(* IEC 61131-3 sources: ia2/library/process-control/pous (part 2) *)

(* ---- fb_pid_3step.st ---- *)
(*
  FB_PID_3STEP — step (3-step) PID: open/close pulse control of a motorized actuator,
  supporting both no-position-feedback (travel-time integral estimate) and
  with-feedback wiring.

  ~ Standard step PID / 3-step output controller (step controller / 3-step PID, driving
  integrating-type actuators such as motorized control valves and motorized dampers),
  found in every major DCS/PLC standard library.

  Purpose: closed-loop control of a motorized actuator (motorized valve / motorized
  damper, which is itself an integrating element: energized it runs open/close, de-energized
  it stops in place). Without a position transmitter, estimate position by integrating
  travel time (pos_fb < 0); with a 4-20 mA position feedback, use it directly.

  Behavior:
    1) Position estimate pos_est: pos_fb >= 0 takes the feedback directly (clamped
       0..100); otherwise integrate from the previous scan's output and the travel time:
       an open pulse adds +100*dt_s/motor_time_s, a close pulse decrements likewise
       (clamped 0..100).
    2) An internal positional PID (reverse-acting e = sp - pv, D on PV with automatic
       3*dt_s PT1 filtering) computes the target position target 0..100; integral
       back-calculation anti-windup; in manual, target tracks pos_est so the return to
       auto is bumpless. For direct-acting scenarios, invert pv/sp externally.
    3) Three-step output: position deviation = target - pos_est;
       > deadband_pct emits an open pulse, < -deadband_pct emits a close pulse, within
       the deadband stop. In auto, once a pulse is emitted it is held at least
       min_pulse_s (to avoid short pulses hammering the contactor); manual jogs
       man_open/man_close pass through (no minimum pulse width, mutually interlocked
       when both are commanded), constrained only by the travel limits. A reversal must
       pass through one scan fully stopped (stop before reversing). At a travel boundary
       (pos_est reaching 0 or 100), stop that direction's pulse immediately.
    Tuning tip: deadband_pct should be larger than the travel corresponding to the
    minimum pulse width (min_pulse_s / motor_time_s * 100%), otherwise it will still
    overshoot and oscillate within the deadband.

  Inputs:
    pv           REAL  process value
    sp           REAL  setpoint
    kp           REAL  proportional gain
    ti_s         REAL  integral time s (0 = no integral)
    td_s         REAL  derivative time s (0 = derivative off)
    dt_s         REAL  sample period s (<= 0 holds this scan, no action)
    motor_time_s REAL  actuator full-travel time s (0->100%; used for estimation and limits)
    min_pulse_s  REAL  minimum pulse width in auto s
    deadband_pct REAL  position deadband % (no action within the deviation deadband)
    auto         BOOL  TRUE auto / FALSE manual jog
    man_open     BOOL  manual open jog (interlocked, no action when commanded with man_close)
    man_close    BOOL  manual close jog
    pos_fb       REAL  position feedback 0..100 % (< 0 = no feedback, use travel estimate)
  Outputs:
    q_open  BOOL  open-direction pulse output
    q_close BOOL  close-direction pulse output
    pos_est REAL  position estimate/feedback 0..100 %
*)
FUNCTION_BLOCK FB_PID_3STEP
  VAR_INPUT
    pv           : REAL;
    sp           : REAL;
    kp           : REAL := 1.0;
    ti_s         : REAL := 0.0;
    td_s         : REAL := 0.0;
    dt_s         : REAL := 0.1;
    motor_time_s : REAL := 60.0;
    min_pulse_s  : REAL := 0.5;
    deadband_pct : REAL := 1.0;
    auto         : BOOL := TRUE;
    man_open     : BOOL := FALSE;
    man_close    : BOOL := FALSE;
    pos_fb       : REAL := -1.0;
  END_VAR
  VAR_OUTPUT
    q_open  : BOOL;
    q_close : BOOL;
    pos_est : REAL;
  END_VAR
  VAR
    i_acc     : REAL; (* positional-PID integral term (back-calculation bumpless) *)
    pv_f      : REAL; (* D-term PT1 filter state *)
    pv_f_prev : REAL;
    t_f       : REAL;
    e         : REAL;
    p_term    : REAL;
    d_term    : REAL;
    target    : REAL; (* PID target position 0..100 *)
    err_pos   : REAL; (* position deviation target - pos_est *)
    pulse_t   : REAL; (* elapsed duration of the current pulse s *)
    open_req  : BOOL; (* open-direction demand this scan *)
    close_req : BOOL;
    init_done : BOOL; (* filter-state first-scan alignment flag *)
  END_VAR

  IF dt_s <= 0.0 THEN
    RETURN; (* invalid sample period: hold *)
  END_IF;

  IF NOT init_done THEN
    pv_f := pv;
    pv_f_prev := pv;
    init_done := TRUE;
  END_IF;

  (* 1) Position estimate: use feedback directly when available; otherwise integrate from the previous scan's output over the travel time *)
  IF pos_fb >= 0.0 THEN
    pos_est := pos_fb;
  ELSE
    IF motor_time_s > 0.0 THEN
      IF q_open THEN
        pos_est := pos_est + 100.0 * dt_s / motor_time_s;
      END_IF;
      IF q_close THEN
        pos_est := pos_est - 100.0 * dt_s / motor_time_s;
      END_IF;
    END_IF;
  END_IF;
  IF pos_est > 100.0 THEN
    pos_est := 100.0;
  ELSIF pos_est < 0.0 THEN
    pos_est := 0.0;
  END_IF;

  (* 2) Positional PID -> target position (reverse-acting; D on PV, automatic 3*dt_s filtering) *)
  t_f := 3.0 * dt_s;
  pv_f := pv_f + dt_s / (t_f + dt_s) * (pv - pv_f);
  e := sp - pv;
  p_term := kp * e;
  d_term := 0.0;
  IF td_s > 0.0 THEN
    d_term := 0.0 - kp * td_s * (pv_f - pv_f_prev) / dt_s;
  END_IF;
  pv_f_prev := pv_f;

  IF auto THEN
    IF ti_s > 0.0 THEN
      i_acc := i_acc + kp * dt_s / ti_s * e;
    END_IF;
    target := p_term + i_acc + d_term;
  ELSE
    target := pos_est; (* Manual: target tracks the current position, bumpless return to auto *)
  END_IF;
  IF target > 100.0 THEN
    target := 100.0;
  ELSIF target < 0.0 THEN
    target := 0.0;
  END_IF;
  IF ti_s > 0.0 OR NOT auto THEN
    i_acc := target - p_term - d_term; (* Back-calculation: anti-windup + bumpless *)
  END_IF;

  (* 3) Three-step output demand *)
  IF auto THEN
    err_pos := target - pos_est;
    open_req := err_pos > deadband_pct;
    close_req := err_pos < 0.0 - deadband_pct;
  ELSE
    open_req := man_open AND NOT man_close; (* Manual jog passes through, interlocked when both commanded *)
    close_req := man_close AND NOT man_open;
  END_IF;

  (* Travel limits: at a boundary, stop emitting that direction's pulse (same in manual/auto) *)
  IF pos_est >= 100.0 THEN
    open_req := FALSE;
  END_IF;
  IF pos_est <= 0.0 THEN
    close_req := FALSE;
  END_IF;

  (* Pulse timing and output: in auto, dropping the demand must satisfy the minimum
     pulse width; in manual, dropping stops immediately; a reversal must pass through
     one scan fully stopped (the current direction drops first, the reverse is allowed
     only on the next scan) *)
  IF q_open OR q_close THEN
    pulse_t := pulse_t + dt_s;
  END_IF;

  IF q_open THEN
    IF pos_est >= 100.0 THEN
      q_open := FALSE; (* at limit, stop *)
    ELSIF NOT open_req AND (NOT auto OR pulse_t >= min_pulse_s) THEN
      q_open := FALSE;
    END_IF;
  ELSIF q_close THEN
    IF pos_est <= 0.0 THEN
      q_close := FALSE;
    ELSIF NOT close_req AND (NOT auto OR pulse_t >= min_pulse_s) THEN
      q_close := FALSE;
    END_IF;
  ELSE
    pulse_t := 0.0;
    IF open_req THEN
      q_open := TRUE;
    ELSIF close_req THEN
      q_close := TRUE;
    END_IF;
  END_IF;
END_FUNCTION_BLOCK

(* ---- fb_pid_pos.st ---- *)
(*
  FB_PID_POS — positional (absolute-output) PID controller with observable p/i/d terms,
  SP weighting, derivative-on-PV (D on PV + PT1 filter), back-calculation anti-windup
  and bumpless transfer.

  ~ Standard positional PID (absolute-output form, observable P/I/D terms, SP weighting
  b, derivative acting on PV), found in every major DCS/PLC standard library.

  Purpose: complements the velocity-form FB_PID -- for loops that need to observe/debug
  the integral term, want SP weighting (b < 1 suppresses the proportional kick on a
  setpoint step), or need an absolute-quantity output downstream. For incremental
  output / cascade relay scenarios, FB_PID is still recommended.

  Algorithm (positional):
    e   := sp - pv (reverse-acting, default); direct = TRUE gives e := pv - sp
    e_p := b*sp - pv (the SP-weighted deviation used only by the P term; reversed when direct)
    p_part := kp * e_p
    i_part := i_part + kp*dt_s/ti_s * e (accumulated when ti_s > 0)
    d_part := -kp*td_s * d(pv_f)/dt (derivative acts on PV: no kick on an SP step;
              pv first passes a PT1 filter, t_dfilt_s <= 0 takes 3*dt_s automatically;
              sign goes positive when direct)
    out := p_part + i_part + d_part + ff, clamped to [out_min, out_max]
  Anti-windup and bumpless (back-calculation): each scan wraps up by back-calculating i_part as
    i_part := out - p_part - d_part - ff
  -- on clamping the integral is pulled back (no windup); in manual/track the output
  follows the supplied value and i_part back-calculates in step, so the return to auto
  has no jump. When ti_s = 0 (no integral), i_part is back-calculated only during
  manual/track (where it is a fixed bias / manual-reset term, not overwritten by
  clamping events during auto, keeping the offset characteristic of P-type control
  stable).
  Mode priority: track > NOT auto (manual) > auto (same as FB_PID).
  Identity: in every mode out = p_part + i_part + d_part + ff (after clamping, except
  on an auto clamping scan with ti_s = 0) -- the sum of the terms is the output,
  intuitive for debugging.

  Inputs:
    pv          REAL  process value
    sp          REAL  setpoint
    kp          REAL  proportional gain
    ti_s        REAL  integral time s (0 = no integral)
    td_s        REAL  derivative time s (0 = derivative off)
    t_dfilt_s   REAL  derivative pre-filter PT1 time constant s (<= 0 = auto 3*dt_s)
    sp_weight_b REAL  SP weighting coefficient b (acts on the P term only; 1 = no weighting,
                      0 = the P term sees pv only -- an SP step gives no proportional kick at all)
    dt_s        REAL  sample period s (<= 0 holds this scan, no action)
    direct      BOOL  TRUE = direct-acting (pv up -> out up), FALSE = reverse-acting
    auto        BOOL  TRUE auto / FALSE manual
    manual_out  REAL  manual output value
    out_min     REAL  output low limit (assumes out_min < out_max)
    out_max     REAL  output high limit
    ff          REAL  feedforward (added to output before clamp)
    track       BOOL  output-tracking enable (highest priority)
    track_value REAL  tracking value
  Outputs:
    out    REAL  control output (clamped in every mode)
    dev    REAL  deviation (reverse-acting sp-pv / direct-acting pv-sp, without SP weighting)
    p_part REAL  proportional term (includes SP weighting)
    i_part REAL  integral term (includes back-calculation correction)
    d_part REAL  derivative term
*)
FUNCTION_BLOCK FB_PID_POS
  VAR_INPUT
    pv          : REAL;
    sp          : REAL;
    kp          : REAL := 1.0;
    ti_s        : REAL := 0.0;
    td_s        : REAL := 0.0;
    t_dfilt_s   : REAL := 0.0;
    sp_weight_b : REAL := 1.0;
    dt_s        : REAL := 0.1;
    direct      : BOOL := FALSE;
    auto        : BOOL := TRUE;
    manual_out  : REAL := 0.0;
    out_min     : REAL := 0.0;
    out_max     : REAL := 100.0;
    ff          : REAL := 0.0;
    track       : BOOL := FALSE;
    track_value : REAL := 0.0;
  END_VAR
  VAR_OUTPUT
    out    : REAL;
    dev    : REAL;
    p_part : REAL;
    i_part : REAL;
    d_part : REAL;
  END_VAR
  VAR
    pv_f      : REAL; (* PV after the D-term PT1 filter *)
    pv_f_prev : REAL; (* previous-scan filtered value, for the backward difference *)
    t_f       : REAL; (* filter time constant actually used *)
    d_pv      : REAL; (* rate of change of the filtered PV, units/s *)
    e         : REAL; (* control deviation (includes the action direction) *)
    e_p       : REAL; (* P-term deviation (SP weighting b) *)
    init_done : BOOL; (* filter-state first-scan alignment flag *)
  END_VAR

  IF dt_s <= 0.0 THEN
    RETURN; (* invalid sample period: hold output and history unchanged *)
  END_IF;

  IF NOT init_done THEN
    pv_f := pv; (* align the filter state: no spurious startup derivative *)
    pv_f_prev := pv;
    init_done := TRUE;
  END_IF;

  (* D-term pre-filter PT1 + backward difference (same core as FB_DERIV) *)
  t_f := t_dfilt_s;
  IF t_f <= 0.0 THEN
    t_f := 3.0 * dt_s;
  END_IF;
  pv_f := pv_f + dt_s / (t_f + dt_s) * (pv - pv_f);
  d_pv := (pv_f - pv_f_prev) / dt_s;
  pv_f_prev := pv_f;

  (* Deviation (by action direction) and the SP-weighted P deviation *)
  IF direct THEN
    e := pv - sp;
    e_p := pv - sp_weight_b * sp;
  ELSE
    e := sp - pv;
    e_p := sp_weight_b * sp - pv;
  END_IF;
  dev := e;

  p_part := kp * e_p;

  d_part := 0.0;
  IF td_s > 0.0 THEN
    (* Derivative acts on PV (no kick on an SP step): reverse-acting, rising pv should push the output down -> negative sign *)
    IF direct THEN
      d_part := kp * td_s * d_pv;
    ELSE
      d_part := 0.0 - kp * td_s * d_pv;
    END_IF;
  END_IF;

  IF track THEN
    (* Output tracking: follows track_value unconditionally, highest priority *)
    out := track_value;
  ELSIF NOT auto THEN
    (* Manual: follows manual_out; the i_part back-calculation guarantees a bumpless return to auto *)
    out := manual_out;
  ELSE
    IF ti_s > 0.0 THEN
      i_part := i_part + kp * dt_s / ti_s * e;
    END_IF;
    out := p_part + i_part + d_part + ff;
  END_IF;

  (* Output clamp *)
  IF out > out_max THEN
    out := out_max;
  ELSIF out < out_min THEN
    out := out_min;
  END_IF;

  (* Back-calculate i_part: makes P+I+D+ff always equal the clamped output -> clamping
     gives anti-windup and manual/track gives bumpless alignment. When ti_s = 0,
     back-calculate only during manual/track (see header note) *)
  IF ti_s > 0.0 OR track OR NOT auto THEN
    i_part := out - p_part - d_part - ff;
  END_IF;
END_FUNCTION_BLOCK

(* ---- fb_pulser.st ---- *)
(*
  FB_PULSER — periodic pulse generator.

  Purpose: periodic air-cannon / air-hammer silo purging, periodic lubrication, heartbeat output.
  Example: once enabled, output a pulse_len_s-wide pulse every period_s seconds (the pulse comes at the period start).

  Behavior:
    while enabled, the phase phase_s accumulates by dt_s manually; q := TRUE while
    phase_s < pulse_len_s, wrapping at period_s (subtraction wrap, so the long-term
    cadence does not drift).
    NOT enable or invalid parameters (period_s/dt_s <= 0) -> q := FALSE and phase cleared
    (re-enabling starts from the pulse).
    pulse_len_s >= period_s -> q is always TRUE (continuous output by definition).

  Inputs:
    enable      BOOL  enable
    period_s    REAL  pulse period s
    pulse_len_s REAL  pulse width s
    dt_s        REAL  sample period s
  Outputs:
    q BOOL  pulse output
*)
FUNCTION_BLOCK FB_PULSER
  VAR_INPUT
    enable      : BOOL;
    period_s    : REAL := 60.0;
    pulse_len_s : REAL := 1.0;
    dt_s        : REAL := 0.1;
  END_VAR
  VAR_OUTPUT
    q : BOOL;
  END_VAR
  VAR
    phase_s : REAL; (* phase within the period 0..period_s, manual timing in place of TP/TON *)
  END_VAR

  IF NOT enable OR period_s <= 0.0 OR dt_s <= 0.0 THEN
    phase_s := 0.0;
    q := FALSE;
    RETURN;
  END_IF;

  (* Emit the pulse by the current phase first (TRUE immediately on the first enabled period), then advance the phase *)
  q := phase_s < pulse_len_s;

  phase_s := phase_s + dt_s;
  IF phase_s >= period_s THEN
    phase_s := phase_s - period_s; (* subtraction wrap, keeps the long-term cadence *)
  END_IF;
END_FUNCTION_BLOCK

(* ---- fb_pv_hold.st ---- *)
(*
  FB_PV_HOLD — bad-PV hold / substitute.

  ~ Standard bad-value handling block (last-good hold / substitute value, including
  bad-value timeout degradation), the standard line of defense before a measurement
  enters a control loop; every major DCS/PLC input-processing chain has an equivalent
  mechanism.

  Purpose: on transmitter open-circuit/over-range (e.g. FB_SCALE.fault, or the inverse
  of FB_MID3.q_fail used as good), give the downstream loop a controlled PV: hold the
  last good value first to ride out chatter, then on timeout hold/substitute/follow as
  configured, while emitting q_bad/q_timeout for alarming and loop-to-manual logic.

  Behavior:
    good = TRUE: out := u, remember the last good value, clear q_bad/q_timeout, clear
    the bad-value timer.
    good = FALSE: q_bad := TRUE, accumulate the bad-value timer (manual dt_s):
      before timeout_s: out := last good value (short chatter rides through on hold);
      at timeout_s (timeout_s = 0 immediately): q_timeout := TRUE, then by mode:
        mode = 0: keep holding the last good value;
        mode = 1: out := sub_value (substitute value, e.g. a safe-side setting);
        mode = 2: out := u (follow the raw value -- just raise the alarm flag without
                  intervening, downstream handles it).
    When bad on the very first scan, the last good value takes the current u (no better history).
    dt_s <= 0 -> the bad-value timer does not advance (when timeout_s > 0, the hold segment is maintained).

  Inputs:
    u         REAL  input (raw PV)
    good      BOOL  input valid (FALSE = bad value; feed the inverse of a quality bit / open-circuit decision)
    mode      REAL  0 = hold last good value / 1 = substitute value / 2 = follow raw value
    sub_value REAL  substitute value (used by mode = 1)
    timeout_s REAL  bad-value persistence timeout s (0 = act by mode immediately; > 0 hold first)
    dt_s      REAL  sample period s
  Outputs:
    out       REAL  processed PV
    q_bad     BOOL  in bad value (level)
    q_timeout BOOL  bad value has timed out (mode in effect)
*)
FUNCTION_BLOCK FB_PV_HOLD
  VAR_INPUT
    u         : REAL;
    good      : BOOL := TRUE;
    mode      : REAL := 0.0;
    sub_value : REAL := 0.0;
    timeout_s : REAL := 0.0;
    dt_s      : REAL := 0.1;
  END_VAR
  VAR_OUTPUT
    out       : REAL;
    q_bad     : BOOL;
    q_timeout : BOOL;
  END_VAR
  VAR
    last_good : REAL; (* last good value *)
    bad_t     : REAL; (* bad-value accumulated persistence time s *)
    init_done : BOOL; (* first-scan seeding flag *)
  END_VAR

  IF NOT init_done THEN
    last_good := u; (* even when bad on the first scan, take the current u as the held value *)
    init_done := TRUE;
  END_IF;

  IF good THEN
    last_good := u;
    out := u;
    q_bad := FALSE;
    q_timeout := FALSE;
    bad_t := 0.0;
    RETURN;
  END_IF;

  q_bad := TRUE;

  (* Before timeout: hold the last good value (the segment that rides out short chatter) *)
  IF timeout_s > 0.0 THEN
    IF dt_s > 0.0 THEN
      bad_t := bad_t + dt_s;
    END_IF;
    IF bad_t < timeout_s THEN
      out := last_good;
      q_timeout := FALSE;
      RETURN;
    END_IF;
  END_IF;

  (* On timeout (or immediately when timeout_s = 0): act by mode *)
  q_timeout := TRUE;
  IF mode >= 1.5 THEN
    out := u;         (* 2 = follow raw value *)
  ELSIF mode >= 0.5 THEN
    out := sub_value; (* 1 = substitute value *)
  ELSE
    out := last_good; (* 0 = hold last good value *)
  END_IF;
END_FUNCTION_BLOCK

(* ---- fb_pwm.st ---- *)
(*
  FB_PWM — time-proportioning output (0..100% command -> fixed-period duty-cycle on/off).

  ~ Time-proportioning (time-proportioning / PWM): continuous quantity -> periodic
  on/off, the customary form for solid-state-relay / solenoid-valve temperature control.

  Purpose: a PID output driving an on/off actuator via a solid-state relay / solenoid
  valve: electric heaters, steam on/off valves, dosing pumps.
  Behavior:
    Phase accumulator as in FB_PULSER: phase_s accumulates by dt_s, wraps by subtraction
    at period_s (so the long-term cadence does not drift); q := phase_s < on_s.
    on_s := u/100 * period_s (u clamped 0..100 first).
    Minimum on/off times (protecting the contactor/SSR/valve, implemented by clamping the effective duty):
      0 < on_s < min_on_s            -> on_s raised to min_on_s;
      0 < period_s - on_s < min_off_s -> on_s squeezed to period_s - min_off_s
      (the off side has higher priority; if min_on_s + min_off_s > period_s the
      parameters are contradictory and the off side wins -- at the extreme it stays
      permanently off, so do not tune it this way).
    u <= 0 -> off for the whole period; u >= 100 -> on for the whole period (full scale
    is unaffected by the minimum on/off clamp).
    NOT enable or period_s/dt_s <= 0 -> q := FALSE and phase cleared (re-enabling starts
    from the period start, on first then off).
    A change in u takes effect immediately (the comparison threshold within the period
    changes at once, no need to wait for the next period).

  Inputs:
    u         REAL  command 0..100 %
    period_s  REAL  PWM period s
    min_on_s  REAL  minimum on time s (0 = no limit)
    min_off_s REAL  minimum off time s (0 = no limit)
    enable    BOOL  enable
    dt_s      REAL  sample period s
  Outputs:
    q         BOOL  time-proportioning output
*)
FUNCTION_BLOCK FB_PWM
  VAR_INPUT
    u         : REAL;
    period_s  : REAL := 10.0;
    min_on_s  : REAL := 0.0;
    min_off_s : REAL := 0.0;
    enable    : BOOL;
    dt_s      : REAL := 0.1;
  END_VAR
  VAR_OUTPUT
    q : BOOL;
  END_VAR
  VAR
    phase_s : REAL; (* phase within the period, manual timing in place of TP/TON *)
    uc      : REAL;
    on_s    : REAL; (* effective on-duration this scan *)
    off_s   : REAL;
  END_VAR

  IF NOT enable OR period_s <= 0.0 OR dt_s <= 0.0 THEN
    phase_s := 0.0;
    q := FALSE;
    RETURN;
  END_IF;

  uc := u;
  IF uc < 0.0 THEN
    uc := 0.0;
  ELSIF uc > 100.0 THEN
    uc := 100.0;
  END_IF;

  on_s := uc * period_s / 100.0;

  (* Minimum on: raise the effective duty (u=0 unaffected) *)
  IF on_s > 0.0 AND on_s < min_on_s THEN
    on_s := min_on_s;
  END_IF;

  (* Minimum off: lower the effective duty (at u=100, off=0 so it does not trigger, stays permanently on) *)
  off_s := period_s - on_s;
  IF off_s > 0.0 AND off_s < min_off_s THEN
    on_s := period_s - min_off_s;
    IF on_s < 0.0 THEN
      on_s := 0.0;
    END_IF;
  END_IF;

  q := phase_s < on_s;

  phase_s := phase_s + dt_s;
  IF phase_s >= period_s THEN
    phase_s := phase_s - period_s; (* subtraction wrap, keeps the long-term cadence *)
  END_IF;
END_FUNCTION_BLOCK

(* ---- fb_ramp.st ---- *)
(*
  FB_RAMP — setpoint ramp generator (rate-limited approach to a fixed target).

  ~ Standard setpoint ramp generator.

  Purpose: gentle setpoint changes (avoiding step shocks to actuators/process),
  segmented heat-up/pressure-up curves.
  Difference from FB_RATE_LIMIT: this block moves toward a fixed target and reports
  ramping; RATE_LIMIT continuously follows a changing input and only clamps the
  per-second change.

  Behavior:
    out approaches target at rate_up (upward) / rate_dn (downward, supplied positive)
    units per second, and on arrival ramping := FALSE. A rate of 0 means a direct
    step in that direction.
    track level-active: out follows track_value unconditionally and ramping := FALSE;
    after track is released, the ramp continues from the current value toward target
    (the bumpless-startup idiom: track-align to the current process value first, then
    release to start ramping).
    dt_s <= 0 -> hold. Note out initializes to 0: on the first startup scan, prefer
    aligning with track.

  Inputs:
    target      REAL  target value
    rate_up     REAL  upward rate units/s (0 = step)
    rate_dn     REAL  downward rate units/s (supplied positive; 0 = step)
    dt_s        REAL  sample period s
    track       BOOL  tracking enable (level-active)
    track_value REAL  tracking value
  Outputs:
    out     REAL  ramp output
    ramping BOOL  ramp in progress (target not yet reached)
*)
FUNCTION_BLOCK FB_RAMP
  VAR_INPUT
    target      : REAL;
    rate_up     : REAL := 0.0;
    rate_dn     : REAL := 0.0;
    dt_s        : REAL := 0.1;
    track       : BOOL := FALSE;
    track_value : REAL := 0.0;
  END_VAR
  VAR_OUTPUT
    out     : REAL;
    ramping : BOOL;
  END_VAR
  VAR
    delta : REAL;
    step  : REAL;
  END_VAR

  IF track THEN
    out := track_value; (* bumpless: after release the ramp continues from here *)
    ramping := FALSE;
    RETURN;
  END_IF;

  IF dt_s <= 0.0 THEN
    RETURN; (* hold *)
  END_IF;

  delta := target - out;
  IF delta > 0.0 THEN
    step := rate_up * dt_s;
    IF rate_up <= 0.0 OR step >= delta THEN
      out := target; (* rate 0 step / reachable this scan *)
      ramping := FALSE;
    ELSE
      out := out + step;
      ramping := TRUE;
    END_IF;
  ELSIF delta < 0.0 THEN
    step := rate_dn * dt_s;
    IF rate_dn <= 0.0 OR step >= 0.0 - delta THEN
      out := target;
      ramping := FALSE;
    ELSE
      out := out - step;
      ramping := TRUE;
    END_IF;
  ELSE
    ramping := FALSE;
  END_IF;
END_FUNCTION_BLOCK

(* ---- fb_rampsoak8.st ---- *)
(*
  FB_RAMPSOAK8 — 8-segment setpoint programmer (ramp-soak setpoint programmer).

  ~ Standard program-setpoint / curve-setpoint block (ramp-soak / setpoint programmer:
  heat-up curves, heat-treatment curves, batch temperature programs), found in every
  major DCS/PLC and program controller.

  Purpose: generate a setpoint from a segmented "ramp to target + soak" curve, feeding
  the sp input of FB_PID / FB_PID_POS: heat-treatment/curing/reactor heat-up programs,
  startup/shutdown load ramp curves. Segment parameters are scalar-expanded sp1..sp8 /
  ramp1_s..ramp8_s / soak1_s..soak8_s (in this dialect an FB-scope array cannot be
  codegen'd, see README gotcha 7; same as FB_CHAR).

  Behavior:
    Each segment N: sp ramps linearly from the previous segment's level (segment 1 from
    sp_init) over rampN_s to spN (rampN_s <= 0 steps), then soaks for soakN_s
    (soaking = TRUE; soakN_s <= 0 passes immediately). Segment parameters latch on the
    segment-entry scan -- changing parameters while running takes effect on the next segment.
    run level-active: TRUE starts and advances the program; FALSE -> return to the start
    (seg := 0, sp := sp_init, done cleared), and setting TRUE again restarts from segment 1.
    hold level-active: freeze sp and the in-segment timer (advance has no effect during hold).
    advance rising edge: jump to the next segment immediately (continue ramping from the
    current sp, curve continuous); advance in the last segment -> done (or cyclic wrap).
    On the last segment's soak end (n_seg clamped 2..8):
      cyclic = FALSE -> done := TRUE, sp pinned at the last segment's target, seg := 0,
      held until reset or run is withdrawn;
      cyclic = TRUE  -> wrap to segment 1 (continue ramping from the current sp, long-term cycling).
    reset level-active (priority): return to start, same as withdrawing run.
    dt_s <= 0 -> no in-segment advance (start/advance edges still handled).

  Inputs:
    sp1..sp8       REAL  per-segment target values (scalar-expanded)
    ramp1_s..ramp8_s REAL  per-segment ramp times s (<= 0 = step)
    soak1_s..soak8_s REAL  per-segment soak times s (<= 0 = no soak)
    n_seg          REAL  number of segments in use 2..8 (auto-clamped)
    run            BOOL  run (level; withdrawing returns to start)
    hold           BOOL  pause (level; freeze sp and the timer)
    advance        BOOL  jump segment (rising edge)
    reset          BOOL  reset (level, priority)
    cyclic         BOOL  TRUE = wrap to segment 1 and cycle after the last segment completes
    sp_init        REAL  start value (the launch level of the segment-1 ramp)
    dt_s           REAL  sample period s
  Outputs:
    sp      REAL  program setpoint output
    seg     REAL  current segment 1..8 (0 = not running / completed)
    soaking BOOL  soak segment in progress
    done    BOOL  program complete (non-cyclic; held until reset / run withdrawn)
*)
FUNCTION_BLOCK FB_RAMPSOAK8
  VAR_INPUT
    sp1     : REAL := 0.0;
    sp2     : REAL := 0.0;
    sp3     : REAL := 0.0;
    sp4     : REAL := 0.0;
    sp5     : REAL := 0.0;
    sp6     : REAL := 0.0;
    sp7     : REAL := 0.0;
    sp8     : REAL := 0.0;
    ramp1_s : REAL := 0.0;
    ramp2_s : REAL := 0.0;
    ramp3_s : REAL := 0.0;
    ramp4_s : REAL := 0.0;
    ramp5_s : REAL := 0.0;
    ramp6_s : REAL := 0.0;
    ramp7_s : REAL := 0.0;
    ramp8_s : REAL := 0.0;
    soak1_s : REAL := 0.0;
    soak2_s : REAL := 0.0;
    soak3_s : REAL := 0.0;
    soak4_s : REAL := 0.0;
    soak5_s : REAL := 0.0;
    soak6_s : REAL := 0.0;
    soak7_s : REAL := 0.0;
    soak8_s : REAL := 0.0;
    n_seg   : REAL := 2.0;
    run     : BOOL := FALSE;
    hold    : BOOL := FALSE;
    advance : BOOL := FALSE;
    reset   : BOOL := FALSE;
    cyclic  : BOOL := FALSE;
    sp_init : REAL := 0.0;
    dt_s    : REAL := 0.1;
  END_VAR
  VAR_OUTPUT
    sp      : REAL;
    seg     : REAL;
    soaking : BOOL;
    done    : BOOL;
  END_VAR
  VAR
    nn         : REAL; (* clamped segment count 2..8 *)
    elapsed_t  : REAL; (* in-segment phase timer s (ramp/soak each start from 0) *)
    level_from : REAL; (* this segment's ramp launch level *)
    seg_sp     : REAL; (* segment parameters latched on entry *)
    seg_ramp_s : REAL;
    seg_soak_s : REAL;
    enter_seg  : REAL; (* segment number to enter this scan (0 = no entry) *)
    go_next    : BOOL; (* segment complete / jump this scan *)
    adv_edge   : BOOL;
    prev_adv   : BOOL; (* advance rising-edge memory *)
  END_VAR

  IF reset THEN
    seg := 0.0;
    soaking := FALSE;
    done := FALSE;
    sp := sp_init;
    elapsed_t := 0.0;
    prev_adv := advance;
    RETURN;
  END_IF;

  adv_edge := advance AND NOT prev_adv;
  prev_adv := advance;

  IF NOT run THEN
    (* Stopped: return to start; re-running starts from segment 1 *)
    seg := 0.0;
    soaking := FALSE;
    done := FALSE;
    sp := sp_init;
    RETURN;
  END_IF;

  IF done THEN
    RETURN; (* Completion hold: sp pinned at the last segment's target, awaiting reset / run withdrawal *)
  END_IF;

  nn := n_seg;
  IF nn < 2.0 THEN
    nn := 2.0;
  ELSIF nn > 8.0 THEN
    nn := 8.0;
  END_IF;

  enter_seg := 0.0;
  go_next := FALSE;

  IF seg < 0.5 THEN
    (* Start: enter segment 1 from sp_init *)
    sp := sp_init;
    enter_seg := 1.0;
  ELSIF hold THEN
    RETURN; (* Freeze: sp and timer held (advance has no effect during hold) *)
  ELSIF adv_edge THEN
    go_next := TRUE; (* Jump segment: continue from the current sp *)
  ELSE
    IF dt_s <= 0.0 THEN
      RETURN; (* invalid sample period: no in-segment advance *)
    END_IF;
    elapsed_t := elapsed_t + dt_s;
    IF NOT soaking THEN
      (* Ramp phase *)
      IF seg_ramp_s <= 0.0 THEN
        sp := seg_sp; (* step segment *)
        soaking := TRUE;
        elapsed_t := 0.0;
      ELSIF elapsed_t >= seg_ramp_s THEN
        sp := seg_sp;
        soaking := TRUE;
        elapsed_t := elapsed_t - seg_ramp_s; (* carry the cross-phase remainder forward *)
      ELSE
        sp := level_from + (seg_sp - level_from) * elapsed_t / seg_ramp_s;
      END_IF;
    END_IF;
    IF soaking AND elapsed_t >= seg_soak_s THEN
      go_next := TRUE; (* soak ended *)
    END_IF;
  END_IF;

  (* Segment-advance decision: last segment -> complete/wrap; otherwise enter the next segment *)
  IF go_next THEN
    IF seg >= nn - 0.5 THEN
      IF cyclic THEN
        enter_seg := 1.0; (* Wrap: segment 1 continues ramping from the current sp *)
      ELSE
        done := TRUE;
        sp := seg_sp; (* Complete: pin at the last segment's target (an early jump also lands here directly) *)
        seg := 0.0;
        soaking := FALSE;
      END_IF;
    ELSE
      enter_seg := seg + 1.0;
    END_IF;
  END_IF;

  (* Segment entry: latch the segment parameters, ramp launches from the current sp *)
  IF enter_seg > 0.5 THEN
    seg := enter_seg;
    level_from := sp;
    elapsed_t := 0.0;
    soaking := FALSE;
    IF seg <= 1.5 THEN
      seg_sp := sp1;
      seg_ramp_s := ramp1_s;
      seg_soak_s := soak1_s;
    ELSIF seg <= 2.5 THEN
      seg_sp := sp2;
      seg_ramp_s := ramp2_s;
      seg_soak_s := soak2_s;
    ELSIF seg <= 3.5 THEN
      seg_sp := sp3;
      seg_ramp_s := ramp3_s;
      seg_soak_s := soak3_s;
    ELSIF seg <= 4.5 THEN
      seg_sp := sp4;
      seg_ramp_s := ramp4_s;
      seg_soak_s := soak4_s;
    ELSIF seg <= 5.5 THEN
      seg_sp := sp5;
      seg_ramp_s := ramp5_s;
      seg_soak_s := soak5_s;
    ELSIF seg <= 6.5 THEN
      seg_sp := sp6;
      seg_ramp_s := ramp6_s;
      seg_soak_s := soak6_s;
    ELSIF seg <= 7.5 THEN
      seg_sp := sp7;
      seg_ramp_s := ramp7_s;
      seg_soak_s := soak7_s;
    ELSE
      seg_sp := sp8;
      seg_ramp_s := ramp8_s;
      seg_soak_s := soak8_s;
    END_IF;
  END_IF;
END_FUNCTION_BLOCK

(* ---- fb_rate_limit.st ---- *)
(*
  FB_RATE_LIMIT — rate limiter (slope clamp that follows the input).

  ~ Standard rate limiter (velocity/slew limiter).

  Purpose: limit the per-second change of a continuously varying signal: valve-command
  anti-chatter, gentle drive-reference changes, feedforward smoothing.
  Difference from FB_RAMP: this block follows a continuously changing input u (no
  target concept) and only clamps |delta|/s; RAMP moves toward a fixed target.

  Behavior:
    delta := u - out is clamped to +/-rate_s*dt_s and then accumulated: out := out + delta_clamped.
    rate_s <= 0 -> pass-through; dt_s <= 0 -> hold;
    reset or first scan -> out := u (alignment, avoiding a full-speed climb from 0 at startup).

  Inputs:
    u      REAL  input
    rate_s REAL  maximum rate of change |units|/s (0 = pass-through)
    dt_s   REAL  sample period s
    reset  BOOL  reset/align (level-active: out follows u)
  Outputs:
    out    REAL  rate-limited output
*)
FUNCTION_BLOCK FB_RATE_LIMIT
  VAR_INPUT
    u      : REAL;
    rate_s : REAL := 0.0;
    dt_s   : REAL := 0.1;
    reset  : BOOL := FALSE;
  END_VAR
  VAR_OUTPUT
    out : REAL;
  END_VAR
  VAR
    delta     : REAL;
    max_step  : REAL;
    init_done : BOOL;
  END_VAR

  IF reset OR NOT init_done THEN
    out := u;
    init_done := TRUE;
    RETURN;
  END_IF;

  IF rate_s <= 0.0 THEN
    out := u; (* pass-through *)
    RETURN;
  END_IF;

  IF dt_s <= 0.0 THEN
    RETURN; (* hold *)
  END_IF;

  delta := u - out;
  max_step := rate_s * dt_s;
  IF delta > max_step THEN
    delta := max_step;
  ELSIF delta < 0.0 - max_step THEN
    delta := 0.0 - max_step;
  END_IF;
  out := out + delta;
END_FUNCTION_BLOCK

(* ---- fb_ratio.st ---- *)
(*
  FB_RATIO — ratio station (ratio setpoint generator).

  ~ Ratio station: the customary block for proportioning/blending loops, output feeds the downstream PID's sp.

  Purpose: ratio control: the follower flow setpoint = wild (leading) flow * ratio +
  bias, and the sp output feeds the sp input of a downstream FB_PID to form the ratio
  loop.
  Example: a follower stream tracks the leading flow at a 0.85 proportion.

  Formula: sp := clamp(ratio, ratio_min, ratio_max) * wild_flow + bias.
  Note: only ratio is clamped (a safety limit on the operator-adjustable ratio), sp is
  not clamped -- sp's dimension follows wild_flow, and the downstream PID has its own
  output clamp.

  Inputs:
    wild_flow REAL  leading flow (the "wild" flow not controlled by this loop)
    ratio     REAL  ratio
    ratio_min REAL  ratio low limit
    ratio_max REAL  ratio high limit
    bias      REAL  bias (engineering units)
  Outputs:
    sp        REAL  follower-loop setpoint
*)
FUNCTION_BLOCK FB_RATIO
  VAR_INPUT
    wild_flow : REAL;
    ratio     : REAL := 1.0;
    ratio_min : REAL := 0.0;
    ratio_max : REAL := 10.0;
    bias      : REAL := 0.0;
  END_VAR
  VAR_OUTPUT
    sp : REAL;
  END_VAR
  VAR
    ratio_used : REAL;
  END_VAR

  ratio_used := ratio;
  IF ratio_used < ratio_min THEN
    ratio_used := ratio_min;
  ELSIF ratio_used > ratio_max THEN
    ratio_used := ratio_max;
  END_IF;

  sp := ratio_used * wild_flow + bias;
END_FUNCTION_BLOCK

(* ---- fb_runtime.st ---- *)
(*
  FB_RUNTIME — equipment run-hours + start-count statistics.

  ~ Equipment run statistics (accumulated run hours + start count), standard
  maintenance data.

  Purpose: pump/fan wear balancing (feed hours to FB_DUTY2's hours_a/b with alt_mode=1),
  maintenance-due reminders, start/stop frequency statistics.
  Behavior:
    while running is TRUE, hours := hours + dt_s/3600;
    on a running rising edge, starts := starts + 1;
    reset level-active clears both (priority, no accumulation during a reset scan).
    The caller may place the instance under VAR RETAIN for retention across power loss
    (same caveat as FB_TOTALIZER: IA2 retain stores as i32, so the retention precision
    of the REAL hours is limited by this; starts is an integer count and is unaffected).

  Inputs:
    running BOOL  equipment running (feed the run feedback, debounce with FB_DEBOUNCE if needed)
    reset   BOOL  clear (level-active, priority; used after maintenance / pump replacement)
    dt_s    REAL  sample period s
  Outputs:
    hours  REAL  accumulated run hours
    starts DINT  accumulated start count
*)
FUNCTION_BLOCK FB_RUNTIME
  VAR_INPUT
    running : BOOL;
    reset   : BOOL := FALSE;
    dt_s    : REAL := 0.1;
  END_VAR
  VAR_OUTPUT
    hours  : REAL;
    starts : DINT;
  END_VAR
  VAR
    prev_run : BOOL; (* rising-edge memory *)
  END_VAR

  IF reset THEN
    hours := 0.0;
    starts := 0;
  ELSE
    IF running AND NOT prev_run THEN
      starts := starts + 1;
    END_IF;
    IF running AND dt_s > 0.0 THEN
      hours := hours + dt_s / 3600.0;
    END_IF;
  END_IF;
  prev_run := running;
END_FUNCTION_BLOCK

(* ---- fb_scale.st ---- *)
(*
  FB_SCALE — linear span conversion: raw counts -> engineering units, with NE43-style open-circuit flag.

  Purpose: analog input scaling. For example, a 4-20 mA signal sampled as raw
  counts (S7-style 5530..27648) is converted to an engineering value such as
  0..100 % or 0..5 m.

  Formula: out := out_min + (raw - raw_min) * (out_max - out_min) / span
           where span = MAX(raw_max - raw_min, 1e-6) (inline IF, divide-by-zero guard).
  Assumes raw_max > raw_min (forward span).

  Inputs:
    raw      REAL  raw count value (e.g. AI channel raw value)
    raw_min  REAL  raw value at span low (4 mA point)
    raw_max  REAL  raw value at span high (20 mA point)
    out_min  REAL  engineering span low
    out_max  REAL  engineering span high
    clamp    BOOL  TRUE clamps output to [out_min, out_max] (reverse engineering span supported)
  Outputs:
    out      REAL  engineering value
    fault    BOOL  raw value out of range >5% of span (NE43-style open-circuit/over-range flag, not latched)
*)
FUNCTION_BLOCK FB_SCALE
  VAR_INPUT
    raw     : REAL;
    raw_min : REAL := 0.0;
    raw_max : REAL := 27648.0;
    out_min : REAL := 0.0;
    out_max : REAL := 100.0;
    clamp   : BOOL := TRUE;
  END_VAR
  VAR_OUTPUT
    out   : REAL;
    fault : BOOL;
  END_VAR
  VAR
    span   : REAL;
    margin : REAL;
    lo     : REAL;
    hi     : REAL;
  END_VAR

  (* span = MAX(raw_max - raw_min, 1e-6) — inline IF, divide-by-zero guard *)
  span := raw_max - raw_min;
  IF span < 0.000001 THEN
    span := 0.000001;
  END_IF;

  (* NE43-style out-of-range test: more than 5% beyond raw span = open-circuit/fault *)
  margin := 0.05 * span;
  fault := (raw < raw_min - margin) OR (raw > raw_max + margin);

  out := out_min + (raw - raw_min) * (out_max - out_min) / span;

  IF clamp THEN
    IF out_min <= out_max THEN
      lo := out_min;
      hi := out_max;
    ELSE
      lo := out_max;
      hi := out_min;
    END_IF;
    IF out < lo THEN
      out := lo;
    ELSIF out > hi THEN
      out := hi;
    END_IF;
  END_IF;
END_FUNCTION_BLOCK

(* ---- fb_select_hl.st ---- *)
(*
  FB_SELECT_HL — high/low selector (override selection).

  ~ High/low selector (override selector), the customary block for override control.

  Purpose: override control -- two controller outputs taking the higher/lower for a
  shared actuator (e.g. compressor anti-surge override, a pressure-override-temperature
  loop); can also take the higher/lower of dual transmitters.

  Behavior: select_high = TRUE takes the greater, FALSE takes the lesser;
  a_selected indicates the output currently comes from a (on a tie, a is deemed
  selected so the indication does not chatter).

  Inputs:
    a           REAL  channel a (typically the primary controller output)
    b           REAL  channel b (typically the override controller output)
    select_high BOOL  TRUE = high select / FALSE = low select
  Outputs:
    out        REAL  selected value
    a_selected BOOL  TRUE = the output currently comes from a
*)
FUNCTION_BLOCK FB_SELECT_HL
  VAR_INPUT
    a           : REAL;
    b           : REAL;
    select_high : BOOL := TRUE;
  END_VAR
  VAR_OUTPUT
    out        : REAL;
    a_selected : BOOL;
  END_VAR

  IF select_high THEN
    IF a >= b THEN
      out := a;
      a_selected := TRUE;
    ELSE
      out := b;
      a_selected := FALSE;
    END_IF;
  ELSE
    IF a <= b THEN
      out := a;
      a_selected := TRUE;
    ELSE
      out := b;
      a_selected := FALSE;
    END_IF;
  END_IF;
END_FUNCTION_BLOCK

(* ---- fb_split_range.st ---- *)
(*
  FB_SPLIT_RANGE — split-range output: one controller output distributed to two valves at the split point.

  ~ Split range: one control output drives two valves by segment (heating/cooling, large/small valves).

  Purpose: one PID drives two actuators: large/small valves extending the range
  (sequential split range, reverse_b := FALSE), or a heating/cooling or
  feed/reflux complementary split range (reverse_b := TRUE, tuned per the actuator's
  air-to-open/air-to-close action and the PID action direction).

  Behavior (u is clamped 0..100 first, both outputs also clamped 0..100):
    out_a: linear 0->100 for u in [0, split], holds 100 once u >= split.
    out_b: linear 0->100 for u in [split, 100], 0 when u <= split;
           when reverse_b = TRUE, segment B reverses to 100->0 (with the end value held
           outside the segment, i.e. out_b = 100 when u <= split, output continuous with
           no jump).
    Curve sketch (split = 50):
      reverse_b = FALSE (large/small valve sequential split range):
        u:     0 .... 50 .... 100
        out_a: 0 -> 100 | holds 100
        out_b: 0   0    | 0 -> 100
      reverse_b = TRUE (complementary, B fully open first then closing):
        u:     0 .... 50 .... 100
        out_a: 0 -> 100 | holds 100
        out_b: 100 100  | 100 -> 0
    Degenerate: split <= 0 -> segment A has no range (u > 0 means 100); split >= 100 ->
    segment B has no range (acts only once u >= 100). split should be set within (0, 100).

  Inputs:
    u         REAL  controller output 0..100
    split     REAL  split point % (segment B start)
    reverse_b BOOL  TRUE = valve B is reverse-acting within its split segment (100->0)
  Outputs:
    out_a     REAL  valve A opening 0..100
    out_b     REAL  valve B opening 0..100
*)
FUNCTION_BLOCK FB_SPLIT_RANGE
  VAR_INPUT
    u         : REAL;
    split     : REAL := 50.0;
    reverse_b : BOOL := TRUE;
  END_VAR
  VAR_OUTPUT
    out_a : REAL;
    out_b : REAL;
  END_VAR
  VAR
    uc     : REAL; (* clamped input *)
    span_b : REAL;
  END_VAR

  (* Input clamp 0..100 *)
  uc := u;
  IF uc < 0.0 THEN
    uc := 0.0;
  ELSIF uc > 100.0 THEN
    uc := 100.0;
  END_IF;

  (* Valve A: 0->100 for u in [0, split] *)
  IF split > 0.0 THEN
    out_a := uc * 100.0 / split;
  ELSE
    (* Degenerate: A has no split segment *)
    IF uc > 0.0 THEN
      out_a := 100.0;
    ELSE
      out_a := 0.0;
    END_IF;
  END_IF;
  IF out_a < 0.0 THEN
    out_a := 0.0;
  ELSIF out_a > 100.0 THEN
    out_a := 100.0;
  END_IF;

  (* Valve B: 0->100 for u in [split, 100] *)
  span_b := 100.0 - split;
  IF span_b > 0.0 THEN
    out_b := (uc - split) * 100.0 / span_b;
  ELSE
    (* Degenerate: B has no split segment *)
    IF uc >= split THEN
      out_b := 100.0;
    ELSE
      out_b := 0.0;
    END_IF;
  END_IF;
  IF out_b < 0.0 THEN
    out_b := 0.0;
  ELSIF out_b > 100.0 THEN
    out_b := 100.0;
  END_IF;

  (* Segment B reverse action (reverse after clamping, hold the end value outside the segment, output continuous) *)
  IF reverse_b THEN
    out_b := 100.0 - out_b;
  END_IF;
END_FUNCTION_BLOCK

(* ---- fb_sqrt_flow.st ---- *)
(*
  FB_SQRT_FLOW — differential-pressure flow square-root extraction.

  ~ DP-flow square-root extraction + low-flow cutoff, a customary block for DCS analog-signal processing.

  Purpose: orifice/venturi/nozzle DP flow measurement: flow is proportional to the
  square root of differential pressure.
  Formula: flow := flow_max * SQRT(dp_pct / 100.0); dp_pct <= cutoff_pct -> flow := 0.
  Notes:
    cutoff_pct is the low-flow cutoff: in the low-DP region the square-root gain tends
    to infinity and noise is amplified severely, so the convention is to cut to zero.
    Default 6.25% (DP) <-> 25% (flow) cutoff point.
    dp_pct <= 0 is treated as 0; dp_pct > 100 is not clipped (the square-root extension
    beyond range is allowed; clamp on the caller side if a hard limit is needed).
    SQRT() is a built-in of this dialect (verified usable through cs project check including codegen).

  Inputs:
    dp_pct     REAL  differential pressure % (0..100, typically fed from FB_SCALE output)
    flow_max   REAL  flow engineering value at 100% DP
    cutoff_pct REAL  low-flow cutoff threshold % (as a DP percentage)
  Outputs:
    flow       REAL  flow engineering value
*)
FUNCTION_BLOCK FB_SQRT_FLOW
  VAR_INPUT
    dp_pct     : REAL;
    flow_max   : REAL := 100.0;
    cutoff_pct : REAL := 6.25;
  END_VAR
  VAR_OUTPUT
    flow : REAL;
  END_VAR

  IF dp_pct <= cutoff_pct OR dp_pct <= 0.0 THEN
    flow := 0.0; (* low-flow cutoff *)
    RETURN;
  END_IF;

  flow := flow_max * SQRT(dp_pct / 100.0);
END_FUNCTION_BLOCK

(* ---- fb_stats.st ---- *)
(*
  FB_STATS — running statistics: min/max/mean/standard deviation (Welford single-pass recurrence).

  ~ Standard statistics block (min/max/average/standard deviation), found in every
  major platform's standard library; this block uses Welford's single-pass
  recurrence -- no arrays, numerically stable.

  Purpose: quality-data statistics (batch temperature mean/spread), measurement
  noise-level assessment, commissioning-time signal profiling (feed FB_AVG_TIME for
  the time average, feed this block for the full-run distribution).
  Behavior (counted by "sample", not consuming dt_s: each scan with enable TRUE counts as 1 sample):
    Welford recurrence (scalar, single-pass, avoiding the precision disaster of
    subtracting squares of large numbers):
      n := n + 1; delta := u - avg; avg := avg + delta / n;
      m2 := m2 + delta * (u - avg)
    sd := SQRT(m2 / n) -- population standard deviation (divide by n, not n-1):
    process monitoring cares about the spread magnitude, the two are indistinguishable
    at large sample counts, and dividing by n is the most direct form in a single-pass
    recurrence.
    reset level-active: clears and re-seeds on the next enabled sample (vmin/vmax/avg
    take that sample's value).
    Note: n is a REAL count; in single precision, after about 1.6E7 samples (about 19
    days at a 100 ms sample) the +1 stops taking effect and the statistics freeze --
    for long-term running, reset per shift / per day.

  Inputs:
    u      REAL  input sample
    enable BOOL  sampling enable (a FALSE scan counts no sample, outputs hold)
    reset  BOOL  clear (level-active, takes priority; re-seeds on the next enabled sample)
  Outputs:
    vmin REAL  minimum value
    vmax REAL  maximum value
    avg  REAL  arithmetic mean
    sd   REAL  population standard deviation
    n    REAL  samples counted so far
*)
FUNCTION_BLOCK FB_STATS
  VAR_INPUT
    u      : REAL;
    enable : BOOL := TRUE;
    reset  : BOOL := FALSE;
  END_VAR
  VAR_OUTPUT
    vmin : REAL;
    vmax : REAL;
    avg  : REAL;
    sd   : REAL;
    n    : REAL;
  END_VAR
  VAR
    m2     : REAL; (* Welford second-order accumulator sum of (u-avg)*(u-avg') *)
    delta  : REAL;
    delta2 : REAL;
  END_VAR

  IF reset THEN
    n := 0.0;
    avg := 0.0;
    m2 := 0.0;
    sd := 0.0;
    vmin := 0.0;
    vmax := 0.0;
    RETURN;
  END_IF;

  IF NOT enable THEN
    RETURN; (* counts no sample: outputs hold *)
  END_IF;

  IF n <= 0.0 THEN
    (* Seed on the first sample *)
    n := 1.0;
    avg := u;
    m2 := 0.0;
    sd := 0.0;
    vmin := u;
    vmax := u;
    RETURN;
  END_IF;

  n := n + 1.0;
  delta := u - avg;
  avg := avg + delta / n;
  delta2 := u - avg;
  m2 := m2 + delta * delta2;
  sd := SQRT(m2 / n);

  IF u < vmin THEN
    vmin := u;
  END_IF;
  IF u > vmax THEN
    vmax := u;
  END_IF;
END_FUNCTION_BLOCK

(* ---- fb_totalizer.st ---- *)
(*
  FB_TOTALIZER — flow totalizer: m3/h instantaneous flow -> m3 accumulated quantity.

  Purpose: feed-water / feed-flow totalizing, shift/batch metering.
  The caller may place the instance under VAR RETAIN so that total is retained with the
  instance across power loss (IA2 snapshots RETAIN variables to state/retain.json).

  Formula: total := total + flow * dt_s / 3600.0 (reset takes priority, no accumulation during a reset scan).
  Note: a negative flow accumulates as usual (bidirectional metering allowed); dt_s <= 0 does not accumulate.

  Inputs:
    flow  REAL  instantaneous flow m3/h
    dt_s  REAL  sample period s
    reset BOOL  clear the total (level-active, takes priority over accumulation)
  Outputs:
    total REAL  accumulated quantity m3
*)
FUNCTION_BLOCK FB_TOTALIZER
  VAR_INPUT
    flow  : REAL;
    dt_s  : REAL := 0.1;
    reset : BOOL;
  END_VAR
  VAR_OUTPUT
    total : REAL;
  END_VAR

  IF reset THEN
    total := 0.0;
  ELSIF dt_s > 0.0 THEN
    total := total + flow * dt_s / 3600.0;
  END_IF;
END_FUNCTION_BLOCK

(* ---- fb_valve.st ---- *)
(*
  FB_VALVE — on/off valve (two-position valve) control, with travel timeout and dual-limit fault monitoring.

  Purpose: standard wrapper for a pneumatic/electric on/off valve, with ZSO/ZSC
  dual-limit feedback.
  Example: the feed valve must be fully open before the downstream may start; a travel
  timeout flags a stuck valve.

  Behavior:
    1) Fault monitoring:
       - zso and zsc TRUE at once -> limit-switch fault, immediate fault;
       - the commanded position and the limit feedback disagree (open valve without zso /
         close valve without zsc) for travel_timeout_s (manual dt_s accumulation) ->
         travel-timeout fault;
       - external fault fault_in -> fault. All latched; reset requires fault_in
         cleared and the dual-limit contradiction absent.
    2) Command latch: cmd_open sets out_open when remote and fault-free;
       cmd_close or fault resets it (fail-safe-close on fault, close takes priority).
    3) Status word status: 0 closed / 1 traveling / 2 open / 3 faulted.

  Inputs:
    cmd_open         BOOL  open command
    cmd_close        BOOL  close command (priority)
    remote           BOOL  remote permissive (gates open only)
    zso              BOOL  open limit (Zero Switch Open)
    zsc              BOOL  close limit (Zero Switch Closed)
    fault_in         BOOL  external fault input
    reset            BOOL  fault reset
    travel_timeout_s REAL  travel timeout s
    dt_s             REAL  sample period s
  Outputs:
    out_open BOOL  open output (TRUE open / FALSE close)
    fault    BOOL  fault (latched)
    status   INT   0 closed / 1 traveling / 2 open / 3 faulted
*)
FUNCTION_BLOCK FB_VALVE
  VAR_INPUT
    cmd_open         : BOOL;
    cmd_close        : BOOL;
    remote           : BOOL := TRUE;
    zso              : BOOL;
    zsc              : BOOL;
    fault_in         : BOOL;
    reset            : BOOL;
    travel_timeout_s : REAL := 30.0;
    dt_s             : REAL := 0.1;
  END_VAR
  VAR_OUTPUT
    out_open : BOOL;
    fault    : BOOL;
    status   : INT;
  END_VAR
  VAR
    travel_t : REAL; (* not-in-position accumulated time s *)
    in_pos   : BOOL;
  END_VAR

  (* 1) Fault monitoring *)
  IF zso AND zsc THEN
    fault := TRUE; (* both limits active at once: limit-switch fault *)
  END_IF;

  in_pos := (out_open AND zso) OR (NOT out_open AND zsc);
  IF in_pos THEN
    travel_t := 0.0;
  ELSE
    travel_t := travel_t + dt_s;
  END_IF;
  IF travel_timeout_s > 0.0 AND travel_t >= travel_timeout_s THEN
    fault := TRUE; (* travel timeout: stuck valve / lost limit *)
  END_IF;

  IF fault_in THEN
    fault := TRUE;
  END_IF;
  IF reset AND NOT fault_in AND NOT (zso AND zsc) THEN
    fault    := FALSE;
    travel_t := 0.0;
  END_IF;

  (* 2) Command latch (close/fault priority, fail-safe-close) *)
  IF cmd_open AND remote AND NOT fault THEN
    out_open := TRUE;
  END_IF;
  IF cmd_close OR fault THEN
    out_open := FALSE;
  END_IF;

  (* 3) Status word *)
  IF fault THEN
    status := 3;
  ELSIF out_open AND zso THEN
    status := 2;
  ELSIF NOT out_open AND zsc THEN
    status := 0;
  ELSE
    status := 1;
  END_IF;
END_FUNCTION_BLOCK

(* ---- demo_main.st ---- *)
(* ============================================================================
  demo_main — mini carbonation-tower loop demonstration PROGRAM.

  The demo instantiates the process-control function blocks that each live in
  their own sibling file (fb_scale.st, fb_pid.st, fb_alarm_hl.st, ...). It is
  meant to be checked together with them: `cs check pous/*.st` resolves the FB
  types across all the files at once, so no block declaration is repeated here.

  Loop wiring (demonstration; variables can be bound to real channels via iomap.toml):
    lt0101_raw (AI raw counts) -> FB_SCALE -> level_pct (tower level %)
    level_pct / level_sp     -> FB_PID (reverse-acting, legacy-signature call, verifies backward compatibility)
                               -> valve_pct (feed control-valve opening)
    level_pct                -> FB_ALARM_HL -> four-level level alarms + any_alm
    hammer_enable            -> FB_PULSER -> hammer_q (periodic air-cannon purge)
    level_pct                -> FB_HILO_FILL -> fill_open (high-close low-open make-up)
    -- the following are extension loops --
    level HH / open-circuit / tower-temp HH / dual-pump fault -> FB_INTERLOCK8 -> ilk_trip + first-out number
    pump_run_fb_a/b          -> FB_RUNTIME x2 -> dual-pump hours / start counts
    fill_open AND NOT ilk    -> FB_DUTY2 (hour balancing) -> dual make-up pumps duty/standby
    gas_flow (leading flow)  -> FB_RATIO -> milk_sp (lime-milk ratio setpoint)
    milk_flow / milk_sp      -> FB_PID (feedforward ff + SP ramp + interlock track forcing)
                               -> FB_SPLIT_RANGE (sequential split range) -> small/large valve
    -- the following demonstrate the math/dynamics blocks (steam-heating cascade + FOPDT plant simulation) --
    steam_valve -> FB_DEADTIME8(20 s) -> manual PT1(30 s) -> tower temp temp_a
                               (dead time + first-order lag = FOPDT plant simulation)
    temp_a / temp_b / bad point -> FB_MID3 (two good one bad, take the average) -> FB_LIMIT -> voted tower temp
    voted tower temp          -> FB_DERIV -> rate of change degC/s;
                               -> FB_STATS (full-run statistics) + FB_AVG_TIME (60 s tumbling window)
    tower-temp master FB_PID -> FB_CASCADE -> steam-flow slave FB_PID -> steam_valve
                               (when not cascaded the master tracks via track, CAS transfer bumpless)
    master PID deviation dev  -> FB_INTEG (interlock hold, clamped +/-1000) -> deviation integral degC*s
    -- the following demonstrate the 0.3.0 loop/device/signal extension blocks (sections 17~26) --
    voted tower temp + q_fail -> FB_PV_HOLD (bad value held 5 s first then hold/substitute) -> temp_held
    heat-up/soak 4-segment curve -> FB_RAMPSOAK8 -> rs_sp (program setpoint)
    temp_held                -> FB_GAIN_SCHED3 (three-zone parameters + boundary transition)
                               -> FB_PID_POS (program SP + scheduled parameters, observable p/i/d)
                               -> FB_MANSTATION (manual station, balance bumpless) -> heat_out
    temp_held / rs_sp        -> FB_PID_3STEP (motorized-actuator pulse control, for observation)
    agitator fwd/rev buttons  -> FB_MOTOR_REV (reversal interlock 2 s, feedback echo simulation)
    fill_open                -> FB_MOV (motorized make-up valve, 30 s simulated travel, dual limits)
    dose start               -> FB_DOSE (coarse 8 / fine 1.5 units/s simulated flow)
    gas_flow + operating p/t  -> FB_FLOW_COMP (square-root DP pressure/temperature compensation) -> gas_flow_std
  scan_s must match the tasks.toml interval_ms (default 100 ms = 0.1 s).
============================================================================ *)

(* ---------------------------------------------------------------------------
   PROGRAM demo_main — wiring layer
--------------------------------------------------------------------------- *)
PROGRAM demo_main
  VAR
    (* -- field signals (bound via iomap; given initial values for the demo) -- *)
    lt0101_raw    : REAL := 13824.0; (* level transmitter raw counts (4-20mA -> 5530..27648) *)
    level_sp      : REAL := 60.0;    (* level setpoint % *)
    alm_ack       : BOOL := FALSE;   (* alarm acknowledge button *)
    hammer_enable : BOOL := TRUE;    (* air cannon in service *)
    gas_flow      : REAL := 1200.0;  (* inlet gas flow m3/h (leading flow FT0201) *)
    milk_flow     : REAL := 950.0;   (* lime-milk flow m3/h (follower pv, FT0202) *)
    milk_ratio    : REAL := 0.85;    (* lime-milk / inlet-gas ratio *)
    pump_run_fb_a : BOOL := FALSE;   (* lime-milk pump 1 run feedback *)
    pump_run_fb_b : BOOL := FALSE;   (* lime-milk pump 2 run feedback *)
    pump_fault_a  : BOOL := FALSE;   (* pump 1 fault (protection relay / thermal overload) *)
    pump_fault_b  : BOOL := FALSE;   (* pump 2 fault *)
    temp_hh       : BOOL := FALSE;   (* tower temperature high-high (external alarm bit) *)
    ilk_reset     : BOOL := FALSE;   (* interlock reset button *)
    rt_reset      : BOOL := FALSE;   (* run-hours clear (after maintenance) *)

    scan_s : REAL := 0.1; (* sample period s, must match tasks.toml interval_ms *)

    (* -- FB instances -- *)
    scale_lt      : FB_SCALE;
    pid_level     : FB_PID;
    alm_level     : FB_ALARM_HL;
    pulser_hammer : FB_PULSER;
    fill_ctl      : FB_HILO_FILL;
    ilk_tower     : FB_INTERLOCK8;
    rt_pump_a     : FB_RUNTIME;
    rt_pump_b     : FB_RUNTIME;
    duty_pumps    : FB_DUTY2;
    ratio_milk    : FB_RATIO;
    pid_milk      : FB_PID;
    split_milk    : FB_SPLIT_RANGE;

    (* -- output / intermediate variables (bound to AO/DO via iomap) -- *)
    level_pct   : REAL; (* tower level % *)
    lt_fault    : BOOL; (* transmitter open-circuit *)
    valve_pct   : REAL; (* feed control-valve opening % *)
    lv_any_alm  : BOOL; (* any level alarm *)
    hammer_q    : BOOL; (* air-cannon solenoid *)
    fill_open   : BOOL; (* make-up demand (high-close low-open) *)
    ilk_trip    : BOOL; (* tower interlock acted *)
    ilk_first   : INT;  (* interlock first-out channel *)
    pump_cmd_a  : BOOL; (* pump 1 start command *)
    pump_cmd_b  : BOOL; (* pump 2 start command *)
    duty_a      : BOOL; (* current duty pump is pump 1 *)
    milk_sp     : REAL; (* lime-milk flow setpoint after ratioing m3/h *)
    milk_dev    : REAL; (* lime-milk loop working deviation (after the SP ramp) *)
    valve_small : REAL; (* lime-milk small-valve opening % (split segment A, fine trim) *)
    valve_big   : REAL; (* lime-milk large-valve opening % (split segment B, range extension) *)

    (* -- math/dynamics block demo: steam-heating cascade + FOPDT plant simulation (sections 12~16) -- *)
    cas_enable     : BOOL := TRUE;  (* cascade-enable switch *)
    temp_sp        : REAL := 75.0;  (* tower-temperature setpoint degC (cascade master SP) *)
    steam_local_sp : REAL := 800.0; (* operator-given steam-flow local SP kg/h when not cascaded *)
    stats_reset    : BOOL := FALSE; (* statistics / deviation-integral clear button *)

    dly_obj      : FB_DEADTIME8; (* plant dead time 20 s *)
    mid_temp     : FB_MID3;      (* tower-temperature median of three (two good one bad) *)
    lim_temp     : FB_LIMIT;     (* voted tower-temperature limit 0..150 degC *)
    deriv_temp   : FB_DERIV;     (* tower-temperature rate of change *)
    casc_temp    : FB_CASCADE;   (* cascade coupling: master output -> steam SP *)
    pid_tc       : FB_PID;       (* cascade master loop: tower temperature *)
    pid_fc_steam : FB_PID;       (* cascade slave loop: steam flow *)
    integ_dev    : FB_INTEG;     (* master-loop deviation integral *)
    stats_temp   : FB_STATS;     (* tower-temperature full-run statistics *)
    avgt_temp    : FB_AVG_TIME;  (* tower-temperature 60 s tumbling-window average *)

    sim_state     : REAL := 40.0; (* FOPDT plant first-order state (manual PT1 discretization, T = 30 s) *)
    temp_a        : REAL;         (* tower-temperature transmitter 1 degC (plant-simulation output) *)
    temp_b        : REAL;         (* redundant point 2 degC (simulated +0.5 degC bias) *)
    temp_voted    : REAL;         (* tower temperature after voting + limiting degC *)
    temp_roc      : REAL;         (* tower-temperature rate of change degC/s *)
    steam_sp_used : REAL;         (* steam slave-loop working SP kg/h (fed back to slave_sp_now) *)
    steam_flow    : REAL;         (* steam flow pv kg/h (simulated static valve characteristic) *)
    steam_valve   : REAL;         (* steam-valve opening % (slave-loop output) *)
    temp_dev_int  : REAL;         (* tower-temperature deviation integral degC*s *)

    (* -- 0.3.0 extension block demo: program setpoint + positional PID chain, device layer,
          compensation (sections 17~26) -- *)
    rs_run       : BOOL := TRUE;  (* program setpoint run *)
    rs_hold      : BOOL := FALSE; (* program setpoint pause *)
    rs_advance   : BOOL := FALSE; (* program setpoint jump-segment button *)
    batch_reset  : BOOL := FALSE; (* program / batch reset button *)
    msta_auto    : BOOL := TRUE;  (* manual station auto in service *)
    msta_man_out : REAL := 0.0;   (* manual station manual output % *)
    agit_fwd_btn : BOOL := FALSE; (* agitator forward button *)
    agit_rev_btn : BOOL := FALSE; (* agitator reverse button *)
    dose_start   : BOOL := FALSE; (* dose start button *)
    dose_abort   : BOOL := FALSE; (* dose abort button *)

    hold_temp  : FB_PV_HOLD;     (* voted tower-temperature bad-value hold *)
    rs_temp    : FB_RAMPSOAK8;   (* heat-up/soak program setpoint *)
    gsch_temp  : FB_GAIN_SCHED3; (* three-zone gain scheduling *)
    pidp_temp  : FB_PID_POS;     (* positional tower-temperature PID (shadow loop) *)
    msta_temp  : FB_MANSTATION;  (* heating-output manual station *)
    pid3s_temp : FB_PID_3STEP;   (* step PID (motorized actuator, for observation) *)
    mrev_agit  : FB_MOTOR_REV;   (* bidirectional agitator motor *)
    mov_fill   : FB_MOV;         (* motorized make-up valve *)
    dose_lime  : FB_DOSE;        (* limestone batch dosing *)
    comp_gas   : FB_FLOW_COMP;   (* inlet-gas pressure/temperature compensation *)

    temp_held    : REAL;          (* tower temperature after bad-value hold degC *)
    rs_sp        : REAL;          (* program setpoint SP degC *)
    heat_out_pos : REAL;          (* positional PID output % *)
    heat_out     : REAL;          (* final heating output after the manual station % *)
    agit_fb_f    : BOOL;          (* agitator forward feedback (output-echo simulation) *)
    agit_fb_r    : BOOL;          (* agitator reverse feedback *)
    mov_sim_pos  : REAL := 0.0;   (* motorized-valve simulated travel 0..100 % *)
    mov_zso      : BOOL := FALSE; (* motorized-valve open limit (simulated) *)
    mov_zsc      : BOOL := TRUE;  (* motorized-valve close limit (simulated, initially fully closed) *)
    mov_q_open   : BOOL;          (* motorized-valve open output (local copy, gotcha 8) *)
    mov_q_close  : BOOL;          (* motorized-valve close output *)
    dose_flow    : REAL := 0.0;   (* dose simulated flow kg/s *)
    dose_q_coar  : BOOL;          (* coarse-feed valve (local copy, gotcha 8) *)
    dose_q_fine  : BOOL;          (* fine-feed valve *)
    gas_flow_std : REAL;          (* standard-condition inlet-gas flow after compensation m3/h *)
  END_VAR

  (* 1) Span conversion: raw counts -> level % *)
  scale_lt(raw := lt0101_raw, raw_min := 5530.0, raw_max := 27648.0,
           out_min := 0.0, out_max := 100.0, clamp := TRUE);
  level_pct := scale_lt.out;
  lt_fault  := scale_lt.fault;

  (* 2) Four-level level alarm, 2% deadband, 3 s delay *)
  alm_level(pv := level_pct, h_sp := 80.0, l_sp := 20.0,
            hh_sp := 90.0, ll_sp := 10.0,
            deadband := 2.0, delay_s := 3.0, dt_s := scan_s, ack := alm_ack);
  lv_any_alm := alm_level.any_alm;

  (* 3) Level PID (reverse-acting: high level -> close the feed valve); on transmitter
        open-circuit, switch to manual and drop to 0. Note: kept as a legacy-signature
        call -- verifies the backward compatibility after the FB_PID upgrade *)
  pid_level(pv := level_pct, sp := level_sp,
            kp := 2.0, ti_s := 120.0, td_s := 0.0, dt_s := scan_s,
            direct := FALSE, auto := NOT lt_fault, manual_out := 0.0,
            out_min := 0.0, out_max := 100.0);
  valve_pct := pid_level.out;

  (* 4) Air cannon: a 2 s purge every 300 s *)
  pulser_hammer(enable := hammer_enable, period_s := 300.0,
                pulse_len_s := 2.0, dt_s := scan_s);
  hammer_q := pulser_hammer.q;

  (* 5) Make-up demand: below 15% needs water, above 85% stops *)
  fill_ctl(pv := level_pct, h_sp := 85.0, l_sp := 15.0);
  fill_open := fill_ctl.valve_open;

  (* 6) Tower interlock summary + first-out: 1=level HH 2=transmitter open-circuit
        3=tower-temp HH 4=dual-pump fault; 5..8 spare, bypassed *)
  ilk_tower(c1 := alm_level.hh_alm,
            c2 := lt_fault,
            c3 := temp_hh,
            c4 := pump_fault_a AND pump_fault_b,
            enable5 := FALSE, enable6 := FALSE,
            enable7 := FALSE, enable8 := FALSE,
            reset := ilk_reset);
  ilk_trip  := ilk_tower.tripped;
  ilk_first := ilk_tower.first_out;

  (* 7) Dual-pump run statistics (hours feed FB_DUTY2 hour balancing; instances may go in VAR RETAIN) *)
  rt_pump_a(running := pump_run_fb_a, reset := rt_reset, dt_s := scan_s);
  rt_pump_b(running := pump_run_fb_b, reset := rt_reset, dt_s := scan_s);

  (* 8) Dual make-up pumps duty/standby: select duty by hour balancing; on interlock action, withdraw demand and stop all *)
  duty_pumps(demand := fill_open AND NOT ilk_trip, alt_mode := 1,
             run_fb_a := pump_run_fb_a, run_fb_b := pump_run_fb_b,
             fault_a := pump_fault_a, fault_b := pump_fault_b,
             hours_a := rt_pump_a.hours, hours_b := rt_pump_b.hours,
             dt_s := scan_s);
  pump_cmd_a := duty_pumps.cmd_a;
  pump_cmd_b := duty_pumps.cmd_b;
  duty_a     := duty_pumps.duty_is_a;

  (* 9) Ratio station: lime-milk flow setpoint = inlet-gas flow x 0.85 (ratio clamped 0.5..1.2) *)
  ratio_milk(wild_flow := gas_flow, ratio := milk_ratio,
             ratio_min := 0.5, ratio_max := 1.2, bias := 0.0);
  milk_sp := ratio_milk.sp;

  (* 10) Lime-milk flow PID: inlet-gas static feedforward (gain 0.01 -> % opening),
         SP ramp 50 (m3/h)/s to avoid a ratio step, interlock action forces the valve
         closed via track *)
  pid_milk(pv := milk_flow, sp := milk_sp,
           kp := 0.8, ti_s := 30.0, td_s := 0.0, dt_s := scan_s,
           direct := FALSE, auto := TRUE, manual_out := 0.0,
           out_min := 0.0, out_max := 100.0,
           ff := gas_flow * 0.01,
           track := ilk_trip, track_value := 0.0,
           sp_rate := 50.0);
  milk_dev := pid_milk.dev;

  (* 11) Split range: PID output 0..50% drives the small valve for fine trim, 50..100%
         the large valve relays (sequential split range, no reversal) *)
  split_milk(u := pid_milk.out, split := 50.0, reverse_b := FALSE);
  valve_small := split_milk.out_a;
  valve_big   := split_milk.out_b;

  (* 12) FOPDT plant simulation: steam-valve opening (previous scan) -> FB_DEADTIME8 dead
         time 20 s -> manual PT1 (T = 30 s, same core as FB_LAG) -> tower temperature.
         Dead time + first-order lag, these two blocks form the most common
         simulation/tuning plant *)
  dly_obj(u := steam_valve, t_delay_s := 20.0, dt_s := scan_s);
  sim_state := sim_state + scan_s / (30.0 + scan_s) * (dly_obj.out - sim_state);
  temp_a := 40.0 + 0.5 * sim_state; (* 0..100 % valve opening -> 40..90 degC *)
  temp_b := temp_a + 0.5;           (* redundant point 2: demo +0.5 degC bias *)

  (* 13) Median of three: point 3's bad value is excluded (good_c := FALSE) -> two good,
         take the average; good channels differing by > 5 degC raise q_dev *)
  mid_temp(a := temp_a, b := temp_b, c := 0.0,
           good_a := TRUE, good_b := TRUE, good_c := FALSE,
           dev_max := 5.0);

  (* 14) Limit the voted value 0..150 degC + filtered derivative (rate of change degC/s for trend/feedforward) *)
  lim_temp(u := mid_temp.out, lo := 0.0, hi := 150.0);
  temp_voted := lim_temp.out;
  deriv_temp(u := temp_voted, t_filt_s := 2.0, dt_s := scan_s);
  temp_roc := deriv_temp.out;

  (* 15) Cascade: tower-temperature master PID (0..100 %) -> FB_CASCADE maps to steam-flow
         SP (0..2000 kg/h) -> steam-flow slave PID -> steam valve. When not cascaded
         (cas_enable = FALSE) the slave uses its local SP and the master tracks the
         equivalent percentage via track, so CAS transfer is bumpless. slave_sp_now is
         fed the previous scan's working SP (standard wiring) *)
  casc_temp(master_out := pid_tc.out, cas_on := cas_enable,
            sp_min := 0.0, sp_max := 2000.0,
            slave_sp_local := steam_local_sp, slave_sp_now := steam_sp_used);
  steam_sp_used := casc_temp.slave_sp;
  pid_tc(pv := temp_voted, sp := temp_sp,
         kp := 1.5, ti_s := 60.0, td_s := 0.0, dt_s := scan_s,
         direct := FALSE, auto := TRUE, manual_out := 0.0,
         out_min := 0.0, out_max := 100.0,
         track := casc_temp.master_track,
         track_value := casc_temp.master_track_value);
  pid_fc_steam(pv := steam_flow, sp := steam_sp_used,
               kp := 0.5, ti_s := 10.0, td_s := 0.0, dt_s := scan_s,
               direct := FALSE, auto := TRUE, manual_out := 0.0,
               out_min := 0.0, out_max := 100.0);
  steam_valve := pid_fc_steam.out;
  steam_flow := steam_valve * 20.0; (* simulated static valve characteristic: 0..100 % -> 0..2000 kg/h *)

  (* 16) Shared-signal (voted tower temperature) statistics trio + deviation integral:
         full-run min/max/mean/standard deviation, 60 s tumbling-window average;
         master-loop deviation integral degC*s (hold on interlock action, clamped +/-1000) *)
  stats_temp(u := temp_voted, enable := TRUE, reset := stats_reset);
  avgt_temp(u := temp_voted, window_s := 60.0, dt_s := scan_s, reset := stats_reset);
  integ_dev(u := pid_tc.dev, k := 1.0, dt_s := scan_s,
            hold := ilk_trip, reset := stats_reset,
            preset := FALSE, preset_value := 0.0,
            out_min := -1000.0, out_max := 1000.0);
  temp_dev_int := integ_dev.out;

  (* 17) Bad-value hold: when the vote is all bad (q_fail), hold the last good value 5 s
         first, then keep holding (mode 0); q_bad/q_timeout feed alarming and loop-to-manual *)
  hold_temp(u := mid_temp.out, good := NOT mid_temp.q_fail,
            mode := 0.0, sub_value := 60.0, timeout_s := 5.0,
            dt_s := scan_s);
  temp_held := hold_temp.out;

  (* 18) 8-segment program setpoint (using 4 segments): a heat-up/soak/cool-down curve
         starting at 40 degC; hold pauses, advance jumps segment, batch_reset resets *)
  rs_temp(sp1 := 55.0, ramp1_s := 120.0, soak1_s := 60.0,
          sp2 := 70.0, ramp2_s := 180.0, soak2_s := 120.0,
          sp3 := 85.0, ramp3_s := 120.0, soak3_s := 300.0,
          sp4 := 40.0, ramp4_s := 240.0, soak4_s := 0.0,
          n_seg := 4.0, run := rs_run, hold := rs_hold,
          advance := rs_advance, reset := batch_reset,
          cyclic := FALSE, sp_init := 40.0, dt_s := scan_s);
  rs_sp := rs_temp.sp;

  (* 19) Three-zone gain scheduling: output PID parameters by zone of the held tower
         temperature (strong in the low-temp zone, weak in the high-temp zone), with a
         +/-2 degC linear transition at the boundaries (interp) *)
  gsch_temp(u_sched := temp_held, x12 := 55.0, x23 := 75.0,
            hyst := 2.0, interp := TRUE,
            kp1 := 2.0, ti1_s := 90.0, td1_s := 0.0,
            kp2 := 1.5, ti2_s := 60.0, td2_s := 0.0,
            kp3 := 1.0, ti3_s := 45.0, td3_s := 0.0);

  (* 20) Positional PID (shadow tower-temperature loop): program setpoint SP + bad-value-held
         PV + scheduled parameters, observable p/i/d; interlock forces 0 via track *)
  pidp_temp(pv := temp_held, sp := rs_sp,
            kp := gsch_temp.kp_out, ti_s := gsch_temp.ti_out_s,
            td_s := gsch_temp.td_out_s, t_dfilt_s := 2.0,
            sp_weight_b := 1.0, dt_s := scan_s,
            direct := FALSE, auto := TRUE, manual_out := 0.0,
            out_min := 0.0, out_max := 100.0,
            ff := 0.0, track := ilk_trip, track_value := 0.0);
  heat_out_pos := pidp_temp.out;

  (* 21) Manual station: in auto pass through the positional PID output (rate-limited
         20 %/s), in manual set directly; balance gives a bumpless return to auto *)
  msta_temp(auto_in := heat_out_pos, auto := msta_auto,
            manual_out := msta_man_out, bias := 0.0, rate := 20.0,
            out_min := 0.0, out_max := 100.0, balance := TRUE,
            dt_s := scan_s);
  heat_out := msta_temp.out;

  (* 22) Step PID (for observation): the same loop driving a motorized actuator without
         position feedback, full travel 60 s, minimum pulse 0.5 s, deadband 1 %, travel estimate pos_est *)
  pid3s_temp(pv := temp_held, sp := rs_sp,
             kp := 1.5, ti_s := 60.0, td_s := 0.0, dt_s := scan_s,
             motor_time_s := 60.0, min_pulse_s := 0.5,
             deadband_pct := 1.0, auto := TRUE,
             man_open := FALSE, man_close := FALSE, pos_fb := -1.0);

  (* 23) Bidirectional agitator motor: forward/reverse buttons, interlock stop has
         priority, reversal interlock 2 s; feedback uses output-echo simulation (one-scan
         lag, never times out) *)
  mrev_agit(cmd_fwd := agit_fwd_btn, cmd_rev := agit_rev_btn,
            stop := ilk_trip, fb_fwd := agit_fb_f, fb_rev := agit_fb_r,
            fb_timeout_s := 5.0, reversal_delay_s := 2.0,
            reset := ilk_reset, dt_s := scan_s);
  agit_fb_f := mrev_agit.q_fwd; (* simulated feedback: output echo (effective next scan) *)
  agit_fb_r := mrev_agit.q_rev;

  (* 24) Motorized make-up valve: make-up demand opens / withdrawal closes (interlock
         forces close), a 30 s simulated travel drives the dual limits; travel-timeout limit 60 s *)
  mov_fill(cmd_open := fill_open AND NOT ilk_trip,
           cmd_close := NOT fill_open OR ilk_trip,
           cmd_stop := FALSE, zso := mov_zso, zsc := mov_zsc,
           travel_s := 60.0, reset := ilk_reset, dt_s := scan_s);
  mov_q_open  := mov_fill.q_open;  (* copy to a local first, then use as an IF condition (gotcha 8) *)
  mov_q_close := mov_fill.q_close;
  IF mov_q_open THEN
    mov_sim_pos := mov_sim_pos + 100.0 * scan_s / 30.0; (* 30 s full-travel simulation *)
  ELSIF mov_q_close THEN
    mov_sim_pos := mov_sim_pos - 100.0 * scan_s / 30.0;
  END_IF;
  IF mov_sim_pos > 100.0 THEN
    mov_sim_pos := 100.0;
  ELSIF mov_sim_pos < 0.0 THEN
    mov_sim_pos := 0.0;
  END_IF;
  mov_zso := mov_sim_pos >= 100.0;
  mov_zsc := mov_sim_pos <= 0.0;

  (* 25) Batch dosing: target 100 kg, fine stage 15 kg, in-flight 2 kg; simulated flow
         coarse 8 / fine 1.5 kg/s (valve state echoed from the previous scan, with a one-scan lag) *)
  dose_lime(start := dose_start, abort := dose_abort,
            flow := dose_flow, target := 100.0,
            fine_qty := 15.0, inflight := 2.0,
            dt_s := scan_s, reset := batch_reset);
  dose_q_coar := dose_lime.q_coarse; (* copy to a local first, then use as an IF condition (gotcha 8) *)
  dose_q_fine := dose_lime.q_fine;
  dose_flow := 0.0;
  IF dose_q_coar THEN
    dose_flow := 8.0;
  ELSIF dose_q_fine THEN
    dose_flow := 1.5;
  END_IF;

  (* 26) Gas pressure/temperature compensation: correct the inlet-gas flow from operating
         150 kPa(g)/45 degC to design conditions (square-root DP, mode 0) -> standard-condition inlet-gas flow *)
  comp_gas(q_raw := gas_flow, p_gauge_kpa := 150.0, t_c := 45.0,
           p_ref_kpa_abs := 201.325, t_ref_c := 20.0,
           atm_kpa := 101.325, mode := 0.0);
  gas_flow_std := comp_gas.q_comp;
END_PROGRAM
